Fanuc KAREL source: kb00053.KL

-- PROVISIONAL review KL for V940-1; original PC SHA256 92132e311ab85a30a540c52700aef7446f06410acdc406f7582a062ff496c0e2
-- Incomplete behavior may be omitted. Consult companion uncertainty JSON. Do not deploy.
PROGRAM KB00053
%NOLOCKGROUP
BEGIN
  -- V9_ZERO_TABLE_METADATA_HINT layout=0002_ascii; no indexed target words; source/name/runtime held
  -- UNRESOLVED_PC offsets 5-15; opcodes 27,31,75
  -- UNRESOLVED_PC offsets 20-24; opcodes 7F
END KB00053
